(* IEC 61131-3 sources: codesys-ai-industrial-robot-control/plc/src/Types, 17 files *)

(* ---- E_AlarmClass.st ---- *)
// Alarm classes (ISA-18.2 style priorities). Critical -> Abort, Error -> Stop.
{attribute 'qualified_only'}
{attribute 'strict'}
TYPE E_AlarmClass :
(
    Info := 0,
    Warning := 1,
    Error := 2,
    Critical := 3
);
END_TYPE

(* ---- E_AlarmId.st ---- *)
// Every alarm of the cell. Definitions (class, text) are in GVL_AlarmDefs.
{attribute 'qualified_only'}
{attribute 'strict'}
TYPE E_AlarmId :
(
    None := 0,
    EStop := 1,
    DoorOpen := 2,
    BridgeLost := 3,
    AxisGroupError := 4,
    ConveyorError := 5,
    FollowingErrorWarn := 6,
    FollowingErrorFault := 7,
    FeedbackStale := 8,
    VacuumNoGrip := 9,
    VacuumLost := 10,
    PartMissed := 11,
    BinFull := 12,
    VisionMissing := 13,
    DecisionFallback := 14,
    LowConfidence := 15,
    QueueOverflow := 16
);
END_TYPE

(* ---- E_Bin.st ---- *)
// Output bins: one per good part type, then the quality bins.
{attribute 'qualified_only'}
{attribute 'strict'}
TYPE E_Bin :
(
    TypeA := 0,
    TypeB := 1,
    TypeC := 2,
    Rework := 3,
    Scrap := 4,
    Quarantine := 5
);
END_TYPE

(* ---- E_DecisionSource.st ---- *)
// Where a part's quality decision came from.
{attribute 'qualified_only'}
{attribute 'strict'}
TYPE E_DecisionSource :
(
    None := 0,
    Ai := 1,
    Fallback := 2
);
END_TYPE

(* ---- E_PackMLCommand.st ---- *)
// PackML state commands.
{attribute 'qualified_only'}
{attribute 'strict'}
TYPE E_PackMLCommand :
(
    None := 0,
    Reset := 1,
    Start := 2,
    Stop := 3,
    Hold := 4,
    Unhold := 5,
    Suspend := 6,
    Unsuspend := 7,
    Abort := 8,
    Clear := 9,
    Complete := 10
);
END_TYPE

(* ---- E_PackMLMode.st ---- *)
// PackML unit modes used by this cell.
{attribute 'qualified_only'}
{attribute 'strict'}
TYPE E_PackMLMode :
(
    Production := 1,
    Maintenance := 2,
    Manual := 3
);
END_TYPE

(* ---- E_PackMLState.st ---- *)
// PackML unit states, numbered as in ISA-TR88.00.02.
{attribute 'qualified_only'}
{attribute 'strict'}
TYPE E_PackMLState :
(
    Undefined := 0,
    Clearing := 1,
    Stopped := 2,
    Starting := 3,
    Idle := 4,
    Suspended := 5,
    Execute := 6,
    Stopping := 7,
    Aborting := 8,
    Aborted := 9,
    Holding := 10,
    Held := 11,
    Unholding := 12,
    Suspending := 13,
    Unsuspending := 14,
    Resetting := 15,
    Completing := 16,
    Complete := 17
);
END_TYPE

(* ---- E_PartState.st ---- *)
// Life cycle of a tracked part.
{attribute 'qualified_only'}
{attribute 'strict'}
TYPE E_PartState :
(
    Free := 0,
    Captured := 1,
    Identified := 2,
    Decided := 3,
    Scheduled := 4,
    Picked := 5,
    Placed := 6,
    Missed := 7,
    Dropped := 8
);
END_TYPE

(* ---- E_PickStep.st ---- *)
// Steps of FB_PickSequence.
{attribute 'qualified_only'}
{attribute 'strict'}
TYPE E_PickStep :
(
    Idle := 0,
    MoveHome := 1,
    MoveReady := 2,
    WaitPart := 3,
    StartTracking := 4,
    Approach := 5,
    Descend := 6,
    Grip := 7,
    Lift := 8,
    MoveToBin := 9,
    Release := 10,
    Retract := 11,
    Aborting := 12,
    Aborted := 13,
    Error := 14,
    RecoverLift := 15       // after an abort with a part on the cup: straight up first
);
END_TYPE

(* ---- E_Quality.st ---- *)
// Quality disposition of a part (spec section 6.3).
{attribute 'qualified_only'}
{attribute 'strict'}
TYPE E_Quality :
(
    Unknown := 0,
    Ok := 1,
    Rework := 2,
    Scrap := 3
);
END_TYPE

(* ---- E_RobotCmd.st ---- *)
// Commands of FB_Robot (start on a rising edge of xExecute).
{attribute 'qualified_only'}
{attribute 'strict'}
TYPE E_RobotCmd :
(
    None := 0,
    MovePtpAcs := 1,       // point-to-point, target in joint space
    MoveLinMcs := 2,       // linear, target in machine coordinates
    MoveLinPcs1 := 3,      // linear, target in PCS_1 (conveyor tracking frame)
    Stop := 4,             // controlled stop, aborts any motion
    Reset := 5,            // reset axis group errors
    MovePtpMcs := 6        // point-to-point, Cartesian target in machine coordinates
);
END_TYPE

(* ---- ST_Alarm.st ---- *)
// Runtime state of one alarm.
TYPE ST_Alarm :
STRUCT
    eClass : E_AlarmClass;
    xActive : BOOL;
    xAcked : BOOL := TRUE;              // no pending acknowledgement
    tRaised : TIME;
END_STRUCT
END_TYPE

(* ---- ST_AlarmDef.st ---- *)
// Static definition of one alarm.
TYPE ST_AlarmDef :
STRUCT
    eClass : E_AlarmClass;
    sText : STRING(80);
END_STRUCT
END_TYPE

(* ---- ST_CaptureMsg.st ---- *)
// Capture request from the PLC to the bridge. A new request has a new udiSeq.
TYPE ST_CaptureMsg :
STRUCT
    udiSeq : UDINT;
    udiPartId : UDINT;
    lrBeltPos : LREAL;                  // conveyor axis position at the trigger [mm]
END_STRUCT
END_TYPE

(* ---- ST_DecisionMsg.st ---- *)
// Quality decision written by the bridge (THX-02). A new message has a new udiSeq.
TYPE ST_DecisionMsg :
STRUCT
    udiSeq : UDINT;
    udiPartId : UDINT;
    eQuality : E_Quality;
    rQualityProb : REAL;
    xIdentReliable : BOOL;
END_STRUCT
END_TYPE

(* ---- ST_PartRecord.st ---- *)
// One tracked part. Positions are in the belt frame at capture time (mm, degrees).
TYPE ST_PartRecord :
STRUCT
    udiPartId : UDINT;
    lrBeltPosAtCapture : LREAL;         // conveyor axis position when PE1 triggered [mm]
    xVisionValid : BOOL;
    usiClass : USINT;                   // detector class index 0..2
    rConfidence : REAL;                 // detector confidence 0..1
    lrX : LREAL;                        // belt frame X at capture [mm]
    lrY : LREAL;                        // belt frame Y [mm]
    lrTheta : LREAL;                    // orientation about Z [deg]
    eQuality : E_Quality;
    rQualityProb : REAL;                // probability of the chosen quality option
    xIdentReliable : BOOL;
    eDecisionSource : E_DecisionSource;
    eTargetBin : E_Bin;
    eState : E_PartState;
    tCaptured : TIME;                   // TIME() at capture
END_STRUCT
END_TYPE

(* ---- ST_VisionMsg.st ---- *)
// Vision result written by the bridge. A new message has a new udiSeq.
TYPE ST_VisionMsg :
STRUCT
    udiSeq : UDINT;
    udiPartId : UDINT;
    xValid : BOOL;
    usiClass : USINT;
    rConfidence : REAL;
    lrX : LREAL;                        // belt frame [mm]
    lrY : LREAL;                        // belt frame [mm]
    lrTheta : LREAL;                    // [deg]
END_STRUCT
END_TYPE
